INTERFACE I_Logger

METHOD CoolingControlLogger
VAR_INPUT
	iLogger		: I_Cooling;
END_VAR
END_METHOD

METHOD GeneratorLogger
VAR_INPUT
	iLogger		: I_Generator;
END_VAR
END_METHOD

METHOD RoomTempLogger : BOOL
VAR_INPUT
	iLogger			: I_RoomTempControl;
END_VAR
END_METHOD

END_INTERFACE

(* stored: Version 1.1.0.1
   Itf I_Logger: Id {92cddb01-eea6-442d-b63b-21c2366cb85a}
   Method CoolingControlLogger: Id {d94e3267-3e83-4ce0-a58d-38680bfb3a7a}
   Method GeneratorLogger: Id {2e68ee11-4676-4d44-a664-a6c65283ecfb}
   Method RoomTempLogger: Id {20ddc7e7-9977-486b-aa83-88fba53294fc} *)
